{attribute 'qualified_only'}
VAR_GLOBAL
	iOutput1 AT %Q*:BOOL;
	iOutput2 AT %Q*:BOOL;
	iOutput3 AT %Q*:BOOL;
	iOutput4 AT %Q*:BOOL;
	
END_VAR

(* stored: Version 1.1.0.1, ProductVersion 3.1.4024.11
   GVL stdOutputs: Id {df674057-7267-0889-0f77-2ec37ce9cd4b} *)
